Staubli VAL3: MonitorIO.pgx

program MonitorIO()
  local bool l_bStopMove
  local bool l_bToHome
  local bool l_bRestartMove
  local bool l_bErr
begin
  l_bRestartMove=true
  l_bStopMove=false
  do
    call io:getDigIO(io:dInput[9],l_bToHome,l_bErr)
    if l_bToHome and (!l_bRestartMove or l_bStopMove)
      l_bRestartMove=true
      l_bStopMove=false
      restartMove()
    endIf

    if !l_bToHome and !l_bStopMove
      l_bStopMove=true
      stopMove()
    endIf

//    if manual:bJogMove
//      if taskStatus("GoHome")>=0
//        taskKill("GoHome")
//      endIf
//      wait(taskStatus("GoHome")<0)

//      stopMove()
//      resetMotion()
//      rs:_nOmacStat=9
//      taskKill("Monitor")
//      wait(taskStatus("Monitor")<0)
//    endIf
    delay(0)
  until false

end
